// TIA Portal project "Safety" (V21)

(* hardware
DEVICE "PLC_Safety"  S7-1500 station
   slot 0: "Rail_0"  Rack  6ES7 590-1***0-0AA0
   slot 1: "PLC_Safety"  CPU 1516F-3 PN/DP  6ES7 516-3FN02-0AB0  V2.9
      slot 3: "CPU display_1"  6ES7591-1BA00-0AA0
      slot 32768: "PROFINET interface_1"  X1
         slot 32769: "Port_1"  X1 P1
         slot 32770: "Port_2"  X1 P2
      slot 33024: "PROFINET interface_2"  X2
         slot 33025: "Port_1"  X2 P1
      slot 33280: "DP interface_1"  X3
      slot 34817: "Virtual CP interface port_1"  Virtual CP interface port  Virtual CP interface port
   slot 2: "F-DI_Main"  F-DI 16x24V DC  6ES7 526-1BH00-0AB0  V1.0
      slot 1: "F-DI_Main"  F-DI 16x24V DC
   slot 3: "F-DQ_Main"  F-DQ 8x24V DC/2A PPM  6ES7 526-2BF00-0AB0  V1.0
      slot 1: "F-DQ_Main"  F-DQ 8x24V DC/2A PPM
DEVICE "Remote_F"  ET 200SP-Station
   slot 0: "Rack_0"  Rack  6ES5 710-8MAx1
   slot 0: "Remote_F"  IM 155-6 PN/2 HF  6ES7 155-6AU01-0CN0  V4.2
   slot 1: "F-DI_Remote"  F-DI 8x24VDC HF  6ES7 136-6BA01-0CA0  V2.0
      slot 1: "F-DI_Remote"  F-DI 8x24VDC HF
   slot 127: "BA 2xRJ45"  BA 2xRJ45  6ES7 193-6AR00-0AA0  V0.0
      slot 1: "Port_1"  X1 P1R  6ES7 193-6AR00-0AA0  V0.0
      slot 2: "Port_2"  X1 P2R  6ES7 193-6AR00-0AA0  V0.0
DEVICE "PLC_Locked"  S7-1500 station
   slot 0: "Rail_0"  Rack  6ES7 590-1***0-0AA0
   slot 1: "PLC_Locked"  CPU 1516F-3 PN/DP  6ES7 516-3FN02-0AB0  V2.9
      slot 3: "CPU display_1"  6ES7591-1BA00-0AA0
      slot 32768: "PROFINET interface_1"  X1
         slot 32769: "Port_1"  X1 P1
         slot 32770: "Port_2"  X1 P2
      slot 33024: "PROFINET interface_2"  X2
         slot 33025: "Port_1"  X2 P1
      slot 33280: "DP interface_1"  X3
      slot 34817: "Virtual CP interface port_1"  Virtual CP interface port  Virtual CP interface port
*)

// ===== PLC "PLC_Safety"  CPU 1516F-3 PN/DP =====
// protected blocks, not shown: "Enable", "Guard", "GuardSafety", "GuardSafety_DB", "LineSafety", "LineSafety_DB", "SafetyData"

VAR_GLOBAL   // PLC tag table "Safety IO"
   "FI_Start" AT %I0.0 : Bool;   // Start button, fail-safe input
   "FI_Stop" AT %I0.1 : Bool;   // Stop button, fail-safe input
   "FI_DoorClosed" AT %I0.2 : Bool;   // Door switch
   "FI_GuardClosed" AT %I20.0 : Bool;   // Guard door switch on the remote station
   "FQ_Motor" AT %Q10.0 : Bool;   // Motor contactor, fail-safe output
   "FQ_Lamp" AT %Q10.1 : Bool;   // Signal lamp, fail-safe output
END_VAR

VAR_GLOBAL   // PLC tag table "Standard"
   "Running" AT %M10.0 : Bool;   // What the safety program released, for the standard program
END_VAR

ORGANIZATION_BLOCK "Main"   // OB1, SCL, ProgramCycle
TITLE = "Main Program Sweep (Cycle)"
{ S7_Optimized_Access := 'TRUE' }
VERSION : 0.1
   VAR_INPUT
      Initial_Call : Bool;   // Initial call of this OB
      Remanence : Bool;   // =True, if remanent data are available
   END_VAR
BEGIN

    // The standard program only reads what the safety program released.
    "Running" := "SafetyData".released;
END_ORGANIZATION_BLOCK

// ===== PLC "PLC_Locked"  CPU 1516F-3 PN/DP =====
// protected blocks, not shown: "LockedSafety", "LockedSafety_DB"